// Tests for MONETcommon.F_AxisTurn, the turn of an azimuth/derotator target inside the axis limits (#2).
// Also MONETcommon.FB_OffsetRamp (2026-11-11), the other helper of the tracking setpoint: here because no suite slot is free
// (MONETcommonTests README, Things to know).
FUNCTION_BLOCK F_AxisTurn_Tests EXTENDS TcUnit.FB_TestSuite
VAR
END_VAR

Site_Limits_Are_Respected();
Endpoints_Are_Inclusive();
No_Valid_Turn_Gives_FALSE_And_The_Nearest_Turn();
Longest_Track_Time_Wins();
No_Velocity_Takes_The_Nearest_Turn();
Margin_Shortens_The_Track_Time();
Hold_Keeps_The_Turn_And_Stops_At_The_Margin();
OffsetRamp_Step_Is_Ramped();
OffsetRamp_Disabled_Follows_At_Once();
OffsetRamp_Retarget_Keeps_The_Velocity_Continuous();
OffsetRamp_SetValue_Blends_To_The_Target();

// The limits are the measured endpoints of each site, never a literal in the library.
METHOD PRIVATE Site_Limits_Are_Respected
VAR
	fPos	: LREAL;
	bOk		: BOOL;
END_VAR
TEST('Site_Limits_Are_Respected');
// MONETS azimuth: 50 deg with negative velocity used to map to 410 and be clamped to 270 (#2)
bOk := MONETcommon.F_AxisTurn(fTarget := 50.0, fVelocity := -0.01, fCurrent := 50.0, bHold := FALSE, fMin := -274.0, fMax := 270.0, fMargin := 1.0, fTrackTimeCap := 14400.0, fPosition => fPos);
AssertTrue(Condition := bOk, Message := 'MONETS az 50');
AssertEquals_LREAL(Expected := 50.0, Actual := fPos, Delta := 1.0E-9, Message := 'MONETS az 50, position');
bOk := MONETcommon.F_AxisTurn(fTarget := 300.0, fVelocity := -0.01, fCurrent := -60.0, bHold := FALSE, fMin := -274.0, fMax := 270.0, fMargin := 1.0, fTrackTimeCap := 14400.0, fPosition => fPos);
AssertTrue(Condition := bOk, Message := 'MONETS az 300 only fits as -60');
AssertEquals_LREAL(Expected := -60.0, Actual := fPos, Delta := 1.0E-9, Message := 'MONETS az 300 only fits as -60, position');
// MONETS derotator: 370 does not fit below 360
bOk := MONETcommon.F_AxisTurn(fTarget := 370.0, fVelocity := 0.01, fCurrent := 10.0, bHold := FALSE, fMin := -90.0, fMax := 360.0, fMargin := 1.0, fTrackTimeCap := 14400.0, fPosition => fPos);
AssertTrue(Condition := bOk, Message := 'MONETS derotator 370');
AssertEquals_LREAL(Expected := 10.0, Actual := fPos, Delta := 1.0E-9, Message := 'MONETS derotator 370, position');
// MONETN derotator: 330 does not fit below 300
bOk := MONETcommon.F_AxisTurn(fTarget := 330.0, fVelocity := 0.01, fCurrent := -30.0, bHold := FALSE, fMin := -170.0, fMax := 300.0, fMargin := 1.0, fTrackTimeCap := 14400.0, fPosition => fPos);
AssertTrue(Condition := bOk, Message := 'MONETN derotator 330');
AssertEquals_LREAL(Expected := -30.0, Actual := fPos, Delta := 1.0E-9, Message := 'MONETN derotator 330, position');
TEST_FINISHED();
END_METHOD

// A window narrower than two turns, so a target has at most one position.
METHOD PRIVATE Endpoints_Are_Inclusive
VAR
	fPos	: LREAL;
	bOk		: BOOL;
END_VAR
TEST('Endpoints_Are_Inclusive');
bOk := MONETcommon.F_AxisTurn(fTarget := 300.0, fVelocity := 0.0, fCurrent := 100.0, bHold := FALSE, fMin := 0.0, fMax := 300.0, fMargin := 1.0, fTrackTimeCap := 14400.0, fPosition => fPos);
AssertTrue(Condition := bOk, Message := 'exactly fMax');
AssertEquals_LREAL(Expected := 300.0, Actual := fPos, Delta := 1.0E-9, Message := 'exactly fMax, position');
bOk := MONETcommon.F_AxisTurn(fTarget := 0.0, fVelocity := 0.0, fCurrent := 100.0, bHold := FALSE, fMin := 0.0, fMax := 300.0, fMargin := 1.0, fTrackTimeCap := 14400.0, fPosition => fPos);
AssertTrue(Condition := bOk, Message := 'exactly fMin');
AssertEquals_LREAL(Expected := 0.0, Actual := fPos, Delta := 1.0E-9, Message := 'exactly fMin, position');
bOk := MONETcommon.F_AxisTurn(fTarget := 301.0, fVelocity := 0.0, fCurrent := 100.0, bHold := FALSE, fMin := 0.0, fMax := 300.0, fMargin := 1.0, fTrackTimeCap := 14400.0, fPosition => fPos);
AssertFalse(Condition := bOk, Message := '1 deg above fMax');
bOk := MONETcommon.F_AxisTurn(fTarget := -1.0, fVelocity := 0.0, fCurrent := 100.0, bHold := FALSE, fMin := 0.0, fMax := 300.0, fMargin := 1.0, fTrackTimeCap := 14400.0, fPosition => fPos);
AssertFalse(Condition := bOk, Message := '1 deg below fMin');
TEST_FINISHED();
END_METHOD

// The result is not to be used for a move; it is the turn nearest to the axis.
METHOD PRIVATE No_Valid_Turn_Gives_FALSE_And_The_Nearest_Turn
VAR
	fPos	: LREAL;
	bOk		: BOOL;
END_VAR
TEST('No_Valid_Turn_Gives_FALSE_And_The_Nearest_Turn');
bOk := MONETcommon.F_AxisTurn(fTarget := 330.0, fVelocity := 0.0, fCurrent := 100.0, bHold := FALSE, fMin := 0.0, fMax := 300.0, fMargin := 1.0, fTrackTimeCap := 14400.0, fPosition => fPos);
AssertFalse(Condition := bOk, Message := '330 in [0, 300], axis at 100');
AssertEquals_LREAL(Expected := -30.0, Actual := fPos, Delta := 1.0E-9, Message := '330 in [0, 300], axis at 100, position');
bOk := MONETcommon.F_AxisTurn(fTarget := 330.0, fVelocity := 0.0, fCurrent := 290.0, bHold := FALSE, fMin := 0.0, fMax := 300.0, fMargin := 1.0, fTrackTimeCap := 14400.0, fPosition => fPos);
AssertFalse(Condition := bOk, Message := '330 in [0, 300], axis at 290');
AssertEquals_LREAL(Expected := 330.0, Actual := fPos, Delta := 1.0E-9, Message := '330 in [0, 300], axis at 290, position');
TEST_FINISHED();
END_METHOD

// MONETN azimuth [-72, 495]: 300 and -60 both fit. 1 deg margin, 4 h cap.
METHOD PRIVATE Longest_Track_Time_Wins
VAR
	fPos	: LREAL;
	bOk		: BOOL;
END_VAR
TEST('Longest_Track_Time_Wins');
// room 193 deg against 553 deg at 0.1 deg/s: 1930 s against 5530 s, both under the cap
bOk := MONETcommon.F_AxisTurn(fTarget := 300.0, fVelocity := 0.1, fCurrent := 300.0, bHold := FALSE, fMin := -72.0, fMax := 495.0, fMargin := 1.0, fTrackTimeCap := 14400.0, fPosition => fPos);
AssertTrue(Condition := bOk, Message := 'positive velocity, -60 has more room');
AssertEquals_LREAL(Expected := -60.0, Actual := fPos, Delta := 1.0E-9, Message := 'positive velocity, -60 has more room, position');
bOk := MONETcommon.F_AxisTurn(fTarget := 100.0, fVelocity := -0.1, fCurrent := 100.0, bHold := FALSE, fMin := -72.0, fMax := 495.0, fMargin := 1.0, fTrackTimeCap := 14400.0, fPosition => fPos);
AssertTrue(Condition := bOk, Message := 'negative velocity, 460 has more room');
AssertEquals_LREAL(Expected := 460.0, Actual := fPos, Delta := 1.0E-9, Message := 'negative velocity, 460 has more room, position');
// slow target: both reach the 4 h cap, the turn nearest to the axis wins (no 360 deg unwind for nothing)
bOk := MONETcommon.F_AxisTurn(fTarget := 100.0, fVelocity := -0.01, fCurrent := 100.0, bHold := FALSE, fMin := -72.0, fMax := 495.0, fMargin := 1.0, fTrackTimeCap := 14400.0, fPosition => fPos);
AssertTrue(Condition := bOk, Message := 'cap tie, axis at 100');
AssertEquals_LREAL(Expected := 100.0, Actual := fPos, Delta := 1.0E-9, Message := 'cap tie, axis at 100, position');
bOk := MONETcommon.F_AxisTurn(fTarget := 100.0, fVelocity := -0.01, fCurrent := 460.0, bHold := FALSE, fMin := -72.0, fMax := 495.0, fMargin := 1.0, fTrackTimeCap := 14400.0, fPosition => fPos);
AssertTrue(Condition := bOk, Message := 'cap tie, axis at 460');
AssertEquals_LREAL(Expected := 460.0, Actual := fPos, Delta := 1.0E-9, Message := 'cap tie, axis at 460, position');
bOk := MONETcommon.F_AxisTurn(fTarget := 300.0, fVelocity := 0.01, fCurrent := 300.0, bHold := FALSE, fMin := -72.0, fMax := 495.0, fMargin := 1.0, fTrackTimeCap := 14400.0, fPosition => fPos);
AssertTrue(Condition := bOk, Message := 'cap tie, positive velocity');
AssertEquals_LREAL(Expected := 300.0, Actual := fPos, Delta := 1.0E-9, Message := 'cap tie, positive velocity, position');
// without a cap the longest track time wins
bOk := MONETcommon.F_AxisTurn(fTarget := 100.0, fVelocity := -0.01, fCurrent := 100.0, bHold := FALSE, fMin := -72.0, fMax := 495.0, fMargin := 1.0, fTrackTimeCap := 1.0E9, fPosition => fPos);
AssertTrue(Condition := bOk, Message := 'no cap');
AssertEquals_LREAL(Expected := 460.0, Actual := fPos, Delta := 1.0E-9, Message := 'no cap, position');
TEST_FINISHED();
END_METHOD

METHOD PRIVATE No_Velocity_Takes_The_Nearest_Turn
VAR
	fPos	: LREAL;
	bOk		: BOOL;
END_VAR
TEST('No_Velocity_Takes_The_Nearest_Turn');
bOk := MONETcommon.F_AxisTurn(fTarget := 100.0, fVelocity := 0.0, fCurrent := 460.0, bHold := FALSE, fMin := -72.0, fMax := 495.0, fMargin := 1.0, fTrackTimeCap := 14400.0, fPosition => fPos);
AssertTrue(Condition := bOk, Message := 'axis at 460');
AssertEquals_LREAL(Expected := 460.0, Actual := fPos, Delta := 1.0E-9, Message := 'axis at 460, position');
bOk := MONETcommon.F_AxisTurn(fTarget := 100.0, fVelocity := 0.0, fCurrent := 100.0, bHold := FALSE, fMin := -72.0, fMax := 495.0, fMargin := 1.0, fTrackTimeCap := 14400.0, fPosition => fPos);
AssertTrue(Condition := bOk, Message := 'axis at 100');
AssertEquals_LREAL(Expected := 100.0, Actual := fPos, Delta := 1.0E-9, Message := 'axis at 100, position');
TEST_FINISHED();
END_METHOD

// MONETS azimuth [-274, 270]: 269.5 is inside the 1 deg margin at the upper end.
METHOD PRIVATE Margin_Shortens_The_Track_Time
VAR
	fPos	: LREAL;
	bOk		: BOOL;
END_VAR
TEST('Margin_Shortens_The_Track_Time');
bOk := MONETcommon.F_AxisTurn(fTarget := 269.5, fVelocity := 0.1, fCurrent := 269.5, bHold := FALSE, fMin := -274.0, fMax := 270.0, fMargin := 1.0, fTrackTimeCap := 14400.0, fPosition => fPos);
AssertTrue(Condition := bOk, Message := '269.5 moving up: the other turn has more room');
AssertEquals_LREAL(Expected := -90.5, Actual := fPos, Delta := 1.0E-9, Message := '269.5 moving up: the other turn has more room, position');
bOk := MONETcommon.F_AxisTurn(fTarget := 269.5, fVelocity := -0.1, fCurrent := 269.5, bHold := FALSE, fMin := -274.0, fMax := 270.0, fMargin := 1.0, fTrackTimeCap := 14400.0, fPosition => fPos);
AssertTrue(Condition := bOk, Message := '269.5 moving down: this turn has more room');
AssertEquals_LREAL(Expected := 269.5, Actual := fPos, Delta := 1.0E-9, Message := '269.5 moving down: this turn has more room, position');
TEST_FINISHED();
END_METHOD

// Tracking: never re-choose, never jump 360 deg; stop 1 deg before the limit.
METHOD PRIVATE Hold_Keeps_The_Turn_And_Stops_At_The_Margin
VAR
	fPos	: LREAL;
	bOk		: BOOL;
END_VAR
TEST('Hold_Keeps_The_Turn_And_Stops_At_The_Margin');
bOk := MONETcommon.F_AxisTurn(fTarget := 100.0, fVelocity := -0.01, fCurrent := 460.0, bHold := TRUE, fMin := -72.0, fMax := 495.0, fMargin := 1.0, fTrackTimeCap := 14400.0, fPosition => fPos);
AssertTrue(Condition := bOk, Message := 'axis at 460, target 100: stays on 460');
AssertEquals_LREAL(Expected := 460.0, Actual := fPos, Delta := 1.0E-9, Message := 'axis at 460, target 100: stays on 460, position');
bOk := MONETcommon.F_AxisTurn(fTarget := 134.5, fVelocity := 0.01, fCurrent := 494.5, bHold := TRUE, fMin := -72.0, fMax := 495.0, fMargin := 1.0, fTrackTimeCap := 14400.0, fPosition => fPos);
AssertFalse(Condition := bOk, Message := '0.5 deg below fMax moving up: inside the margin');
AssertEquals_LREAL(Expected := 494.5, Actual := fPos, Delta := 1.0E-9, Message := '0.5 deg below fMax moving up: inside the margin, position');
bOk := MONETcommon.F_AxisTurn(fTarget := 133.9, fVelocity := 0.01, fCurrent := 493.9, bHold := TRUE, fMin := -72.0, fMax := 495.0, fMargin := 1.0, fTrackTimeCap := 14400.0, fPosition => fPos);
AssertTrue(Condition := bOk, Message := '1.1 deg below fMax moving up');
AssertEquals_LREAL(Expected := 493.9, Actual := fPos, Delta := 1.0E-9, Message := '1.1 deg below fMax moving up, position');
bOk := MONETcommon.F_AxisTurn(fTarget := 135.2, fVelocity := 0.01, fCurrent := 494.9, bHold := TRUE, fMin := -72.0, fMax := 495.0, fMargin := 1.0, fTrackTimeCap := 14400.0, fPosition => fPos);
AssertFalse(Condition := bOk, Message := 'target past fMax: stop, do not jump back to 135.2');
AssertEquals_LREAL(Expected := 495.2, Actual := fPos, Delta := 1.0E-9, Message := 'target past fMax: stop, do not jump back to 135.2, position');
bOk := MONETcommon.F_AxisTurn(fTarget := 269.5, fVelocity := -0.01, fCurrent := 269.5, bHold := TRUE, fMin := -274.0, fMax := 270.0, fMargin := 1.0, fTrackTimeCap := 14400.0, fPosition => fPos);
AssertTrue(Condition := bOk, Message := 'near fMax but moving away');
AssertEquals_LREAL(Expected := 269.5, Actual := fPos, Delta := 1.0E-9, Message := 'near fMax but moving away, position');
bOk := MONETcommon.F_AxisTurn(fTarget := 270.4, fVelocity := -0.01, fCurrent := -89.5, bHold := TRUE, fMin := -90.0, fMax := 360.0, fMargin := 1.0, fTrackTimeCap := 14400.0, fPosition => fPos);
AssertFalse(Condition := bOk, Message := 'derotator 0.5 deg above fMin moving down');
AssertEquals_LREAL(Expected := -89.6, Actual := fPos, Delta := 1.0E-9, Message := 'derotator 0.5 deg above fMin moving down, position');
TEST_FINISHED();
END_METHOD

// FB_OffsetRamp (MONETN 2026-11-11, plan 2026-11-11-altaz-offset-ramp): a 0.01 deg step of the request (the offset step that
// rang with 64-70 % overshoot on the MONETN elevation) reaches the applied value in about 0.43 s, at most 1.6 arcsec per 10 ms
// scan, the velocity changes by at most about fAcceleration * tCycle per scan (no kick), no overshoot.
METHOD PRIVATE OffsetRamp_Step_Is_Ramped
VAR
	fbRamp		: MONETcommon.FB_OffsetRamp;
	i			: INT;
	nDone		: INT;
	fPrev		: LREAL;
	fVel		: LREAL;
	fPrevVel	: LREAL;
	fMaxStep	: LREAL;
	fMaxDv		: LREAL;
	fMax		: LREAL;
	fFirst		: LREAL;
END_VAR
TEST('OffsetRamp_Step_Is_Ramped');
FOR i := 1 TO 200 DO
	fbRamp(fTarget := 0.01, bEnable := TRUE, fAcceleration := 0.2, fVelocity := 0.5, tCycle := T#10MS);
	IF i = 1 THEN
		fFirst := fbRamp.fValue;
	END_IF
	fVel := (fbRamp.fValue - fPrev) / 0.01;
	fMaxStep := MAX(fMaxStep, ABS(fbRamp.fValue - fPrev));
	fMaxDv := MAX(fMaxDv, ABS(fVel - fPrevVel));
	fMax := MAX(fMax, fbRamp.fValue);
	IF fbRamp.bDone AND nDone = 0 THEN
		nDone := i;
	END_IF
	fPrev := fbRamp.fValue;
	fPrevVel := fVel;
END_FOR
AssertTrue(Condition := fFirst < 0.0001, Message := 'the first scan moves the applied value by far less than the step');
AssertTrue(Condition := fMaxStep < 0.0005, Message := 'at most 0.0005 deg (1.8 arcsec) per scan');
AssertTrue(Condition := fMaxDv < 0.003, Message := 'the velocity changes by at most 0.003 deg/s per scan (a step is 1 deg/s)');
AssertTrue(Condition := fMax <= 0.01 + 1.0E-12, Message := 'no overshoot');
AssertTrue(Condition := nDone >= 30 AND nDone <= 50, Message := 'reaches 0.01 deg after 0.3..0.5 s');
AssertEquals_LREAL(Expected := 0.01, Actual := fbRamp.fValue, Delta := 1.0E-12, Message := 'ends on the target');
AssertEquals_LREAL(Expected := 0.0, Actual := fbRamp.fRate, Delta := 1.0E-12, Message := 'ends at rest');
TEST_FINISHED();
END_METHOD

// FB_OffsetRamp outside a track (bEnable FALSE) and with fAcceleration = 0 (the switch back to the old behaviour): the applied
// value is the request in the same call.
METHOD PRIVATE OffsetRamp_Disabled_Follows_At_Once
VAR
	fbRamp		: MONETcommon.FB_OffsetRamp;
END_VAR
TEST('OffsetRamp_Disabled_Follows_At_Once');
fbRamp(fTarget := 0.01, bEnable := FALSE, fAcceleration := 0.2, fVelocity := 0.5, tCycle := T#10MS);
AssertEquals_LREAL(Expected := 0.01, Actual := fbRamp.fValue, Delta := 1.0E-12, Message := 'disabled: at once');
AssertTrue(Condition := fbRamp.bDone, Message := 'disabled: done');
fbRamp(fTarget := -0.02, bEnable := TRUE, fAcceleration := 0.0, fVelocity := 0.5, tCycle := T#10MS);
AssertEquals_LREAL(Expected := -0.02, Actual := fbRamp.fValue, Delta := 1.0E-12, Message := 'fAcceleration 0: at once');
fbRamp(fTarget := 0.03, bEnable := TRUE, fAcceleration := 0.2, fVelocity := 0.0, tCycle := T#10MS);
AssertEquals_LREAL(Expected := 0.03, Actual := fbRamp.fValue, Delta := 1.0E-12, Message := 'fVelocity 0: at once');
// enabled again at rest on the target: nothing moves
fbRamp(fTarget := 0.03, bEnable := TRUE, fAcceleration := 0.2, fVelocity := 0.5, tCycle := T#10MS);
AssertEquals_LREAL(Expected := 0.03, Actual := fbRamp.fValue, Delta := 1.0E-12, Message := 'enabled on the target: stays');
AssertTrue(Condition := fbRamp.bDone, Message := 'enabled on the target: done');
TEST_FINISHED();
END_METHOD

// FB_OffsetRamp: a new request during a ramp (an MQTT offset, then the opposite one 0.15 s later) is taken from the current value
// and velocity: no velocity step, no overshoot past the new target, ends on it. Also a large offset is capped at fVelocity.
METHOD PRIVATE OffsetRamp_Retarget_Keeps_The_Velocity_Continuous
VAR
	fbRamp		: MONETcommon.FB_OffsetRamp;
	fbBig		: MONETcommon.FB_OffsetRamp;
	i			: INT;
	fPrev		: LREAL;
	fVel		: LREAL;
	fPrevVel	: LREAL;
	fMaxDv		: LREAL;
	fMin		: LREAL;
	fMaxVel		: LREAL;
END_VAR
TEST('OffsetRamp_Retarget_Keeps_The_Velocity_Continuous');
FOR i := 1 TO 300 DO
	fbRamp(fTarget := SEL(i > 15, 0.01, -0.01), bEnable := TRUE, fAcceleration := 0.2, fVelocity := 0.5, tCycle := T#10MS);
	fVel := (fbRamp.fValue - fPrev) / 0.01;
	fMaxDv := MAX(fMaxDv, ABS(fVel - fPrevVel));
	fMin := MIN(fMin, fbRamp.fValue);
	fPrev := fbRamp.fValue;
	fPrevVel := fVel;
END_FOR
AssertTrue(Condition := fMaxDv < 0.003, Message := 'retarget: the velocity changes by at most 0.003 deg/s per scan');
AssertTrue(Condition := fMin >= -0.01 - 1.0E-12, Message := 'retarget: no overshoot past the new target');
AssertEquals_LREAL(Expected := -0.01, Actual := fbRamp.fValue, Delta := 1.0E-12, Message := 'retarget: ends on the new target');
AssertTrue(Condition := fbRamp.bDone, Message := 'retarget: done');
// 2 deg: the velocity is capped at fVelocity
fPrev := 0.0;
FOR i := 1 TO 700 DO
	fbBig(fTarget := 2.0, bEnable := TRUE, fAcceleration := 0.2, fVelocity := 0.5, tCycle := T#10MS);
	fMaxVel := MAX(fMaxVel, ABS(fbBig.fValue - fPrev) / 0.01);
	fPrev := fbBig.fValue;
END_FOR
AssertTrue(Condition := fMaxVel <= 0.5 + 1.0E-9, Message := '2 deg: at most fVelocity');
AssertEquals_LREAL(Expected := 2.0, Actual := fbBig.fValue, Delta := 1.0E-12, Message := '2 deg: ends on the target (6.5 s)');
TEST_FINISHED();
END_METHOD

// FB_OffsetRamp.SetValue, the track-start blend of FB_MonetTelescopeControl: the blend starts at the gap between the axis and
// the target (0.008 deg, the azimuth gap seen on MONETN after a slew into tracking) at rest and ramps it to 0 without crossing it.
METHOD PRIVATE OffsetRamp_SetValue_Blends_To_The_Target
VAR
	fbRamp		: MONETcommon.FB_OffsetRamp;
	i			: INT;
	fMin		: LREAL := 1.0;
	fFirst		: LREAL;
END_VAR
TEST('OffsetRamp_SetValue_Blends_To_The_Target');
fbRamp.SetValue(0.008);
AssertEquals_LREAL(Expected := 0.008, Actual := fbRamp.fValue, Delta := 1.0E-12, Message := 'SetValue: the value at once');
AssertFalse(Condition := fbRamp.bDone, Message := 'SetValue: not done');
FOR i := 1 TO 100 DO
	fbRamp(fTarget := 0.0, bEnable := TRUE, fAcceleration := 0.2, fVelocity := 0.5, tCycle := T#10MS);
	IF i = 1 THEN
		fFirst := fbRamp.fValue;
	END_IF
	fMin := MIN(fMin, fbRamp.fValue);
END_FOR
AssertTrue(Condition := ABS(fFirst - 0.008) < 0.0001, Message := 'the first blend scan stays next to the axis position');
AssertTrue(Condition := fMin >= -1.0E-12, Message := 'the blend does not cross the target');
AssertEquals_LREAL(Expected := 0.0, Actual := fbRamp.fValue, Delta := 1.0E-12, Message := 'blended out within 1 s');
TEST_FINISHED();
END_METHOD

END_FUNCTION_BLOCK

(* stored: Version 1.1.0.1, ProductVersion 3.1.4024.15
   POU F_AxisTurn_Tests: Id {6cff4d78-8be6-449c-b836-63b1f5df27f9}, SpecialFunc None
   Method Site_Limits_Are_Respected: Id {edd1381d-aa53-4055-8b95-4c2117652a2c}
   Method Endpoints_Are_Inclusive: Id {6349fddd-f404-4d53-bc63-d26d10284475}
   Method No_Valid_Turn_Gives_FALSE_And_The_Nearest_Turn: Id {0cea74a2-56ad-43ed-ad38-cbf4f58fad34}
   Method Longest_Track_Time_Wins: Id {c3a57a23-db25-41d4-b637-e851b3b9365c}
   Method No_Velocity_Takes_The_Nearest_Turn: Id {61de08ef-e0c3-4a88-976c-94ac3c1ce7a0}
   Method Margin_Shortens_The_Track_Time: Id {5d08f88f-4064-41cd-a630-bdffe4dedb34}
   Method Hold_Keeps_The_Turn_And_Stops_At_The_Margin: Id {6b460c25-f83d-4de3-a448-d37ba4122452}
   Method OffsetRamp_Step_Is_Ramped: Id {5ecf93ab-46f8-4714-bd71-57c68eef0403}
   Method OffsetRamp_Disabled_Follows_At_Once: Id {75829b9a-90df-4d21-93bf-8b717635c8df}
   Method OffsetRamp_Retarget_Keeps_The_Velocity_Continuous: Id {762aebe9-ead3-425a-a79a-12f5a73c19ae}
   Method OffsetRamp_SetValue_Blends_To_The_Target: Id {f73c607f-f2f9-4c70-a5ed-349ec377a4b5} *)
